DATA_BLOCK "DB LAUER"
TITLE =
VERSION : 0.0


  STRUCT
   D_0 : WORD ;
   D_1 : WORD ;
   D_2 : WORD ;
   D_3 : WORD  := W#16#A1;
   D_4 : WORD ;
   D_5 : WORD ;
   D_6 : WORD ;
   D_7 : WORD ;
   D_8 : WORD ;
   D_9 : WORD  := W#16#2006;
   D_10 : WORD  := W#16#1023;
   D_11 : WORD  := W#16#13;
   D_12 : WORD  := W#16#3439;
   D_13 : WORD  := W#16#3500;
   D_14 : WORD ;
   D_15 : WORD  := W#16#1A0;
   D_16 : WORD ;
   D_17 : WORD ;
   D_18 : WORD  := W#16#7C02;
   D_19 : WORD ;
   D_20 : WORD ;
   D_21 : WORD ;
   D_22 : WORD ;
   D_23 : WORD ;
   D_24 : WORD  := W#16#8480;
   D_25 : WORD ;
   D_26 : WORD ;
   D_27 : WORD ;
   D_28 : WORD ;
   D_29 : WORD ;
   D_30 : WORD ;
   D_31 : WORD ;
   D_32 : WORD ;
   D_33 : WORD ;
   D_34 : WORD ;
   D_35 : WORD ;
   D_36 : WORD  := W#16#F00;
   D_37 : WORD  := W#16#3001;
   D_38 : WORD ;
   D_39 : WORD ;
   D_40 : WORD ;
   D_41 : WORD ;
   D_42 : WORD ;
   D_43 : WORD ;
   D_44 : WORD ;
   D_45 : WORD ;
   D_46 : WORD ;
   D_47 : WORD ;
   D_48 : WORD ;
   D_49 : WORD ;
   D_50 : WORD ;
   D_51 : WORD ;
   D_52 : WORD ;
   D_53 : WORD ;
   D_54 : WORD ;
   D_55 : WORD ;
   D_56 : WORD ;
   D_57 : WORD ;
   D_58 : WORD ;
   D_59 : WORD ;
   D_60 : WORD ;
   D_61 : WORD ;
   D_62 : WORD ;
   D_63 : WORD ;
   D_64 : WORD ;
   D_65 : WORD ;
   D_66 : WORD ;
   D_67 : WORD ;
   D_68 : WORD ;
   D_69 : WORD ;
   D_70 : WORD ;
   D_71 : WORD ;
   D_72 : WORD ;
   D_73 : WORD ;
   D_74 : WORD ;
   D_75 : WORD ;
   D_76 : WORD ;
   D_77 : WORD  := W#16#4;
   D_78 : WORD  := W#16#2;
   D_79 : WORD  := W#16#1;
   D_80 : WORD  := W#16#1;
   D_81 : WORD  := W#16#1;
   D_82 : WORD  := W#16#1;
   D_83 : WORD  := W#16#1;
   D_84 : WORD  := W#16#2;
   D_85 : WORD  := W#16#3;
   D_86 : WORD  := W#16#2;
   D_87 : WORD  := W#16#1;
   D_88 : WORD  := W#16#1;
   D_89 : WORD  := W#16#3;
   D_90 : WORD  := W#16#4;
   D_91 : WORD  := W#16#7;
   D_92 : WORD  := W#16#9;
   D_93 : WORD  := W#16#3;
   D_94 : WORD  := W#16#3;
   D_95 : WORD  := W#16#4;
   D_96 : WORD  := W#16#1;
   D_97 : WORD  := W#16#1;
   D_98 : WORD  := W#16#1;
   D_99 : WORD  := W#16#1;
   D_100 : WORD  := W#16#1;
   D_101 : WORD  := W#16#1;
   D_102 : WORD  := W#16#1;
   D_103 : WORD ;
   D_104 : WORD ;
   D_105 : WORD ;
   D_106 : WORD ;
   D_107 : WORD ;
   D_108 : WORD ;
   D_109 : WORD ;
   D_110 : WORD  := W#16#2;
   D_111 : WORD ;
   D_112 : WORD ;
   D_113 : WORD ;
   D_114 : WORD ;
   D_115 : WORD ;
   D_116 : WORD ;
   D_117 : WORD  := W#16#7;
   D_118 : WORD  := W#16#1;
   D_119 : WORD  := W#16#1;
   D_120 : WORD  := W#16#2010;
   D_121 : WORD  := W#16#58;
   D_122 : WORD  := W#16#2010;
   D_123 : WORD  := W#16#2090;
   D_124 : WORD  := W#16#9;
   D_125 : WORD ;
   D_126 : WORD  := W#16#15;
   D_127 : WORD ;
   D_128 : WORD ;
   D_129 : WORD  := W#16#6;
   D_130 : WORD  := W#16#320;
   D_131 : WORD ;
   D_132 : WORD  := W#16#B7;
   D_133 : WORD  := W#16#1EDE;
   D_134 : WORD ;
   D_135 : WORD ;
   D_136 : WORD ;
   D_137 : WORD ;
   D_138 : WORD ;
   D_139 : WORD ;
   D_140 : WORD  := W#16#320;
   D_141 : WORD ;
   D_142 : WORD  := W#16#37;
   D_143 : WORD  := W#16#5D2;
   D_144 : WORD ;
   D_145 : WORD ;
   D_146 : WORD ;
   D_147 : WORD ;
   D_148 : WORD ;
   D_149 : WORD ;
   D_150 : WORD  := W#16#5C;
   D_151 : WORD ;
   D_152 : WORD ;
   D_153 : WORD ;
   D_154 : WORD ;
   D_155 : WORD ;
   D_156 : WORD ;
   D_157 : WORD ;
   D_158 : WORD ;
   D_159 : WORD ;
   D_160 : WORD  := W#16#320;
   D_161 : WORD ;
   D_162 : WORD  := W#16#B9;
   D_163 : WORD  := W#16#181F;
   D_164 : WORD ;
   D_165 : WORD ;
   D_166 : WORD ;
   D_167 : WORD ;
   D_168 : WORD ;
   D_169 : WORD ;
   D_170 : WORD  := W#16#320;
   D_171 : WORD ;
   D_172 : WORD  := W#16#F;
   D_173 : WORD  := W#16#14B9;
   D_174 : WORD ;
   D_175 : WORD ;
   D_176 : WORD ;
   D_177 : WORD ;
   D_178 : WORD ;
   D_179 : WORD ;
   D_180 : WORD  := W#16#320;
   D_181 : WORD ;
   D_182 : WORD ;
   D_183 : WORD  := W#16#4B0;
   D_184 : WORD  := W#16#1;
   D_185 : WORD  := W#16#1;
   D_186 : WORD ;
   D_187 : WORD ;
   D_188 : WORD ;
   D_189 : WORD ;
   D_190 : WORD ;
   D_191 : WORD ;
   D_192 : WORD ;
   D_193 : WORD ;
   D_194 : WORD ;
   D_195 : WORD ;
   D_196 : WORD ;
   D_197 : WORD ;
   D_198 : WORD ;
   D_199 : WORD ;
   D_200 : WORD ;
   D_201 : WORD ;
   D_202 : WORD ;
   D_203 : WORD ;
   D_204 : WORD ;
   D_205 : WORD ;
   D_206 : WORD ;
   D_207 : WORD ;
   D_208 : WORD ;
   D_209 : WORD ;
   D_210 : WORD ;
   D_211 : WORD ;
   D_212 : WORD ;
   D_213 : WORD ;
   D_214 : WORD ;
   D_215 : WORD ;
   D_216 : WORD ;
   D_217 : WORD ;
   D_218 : WORD ;
   D_219 : WORD ;
   D_220 : WORD ;
   D_221 : WORD ;
   D_222 : WORD ;
   D_223 : WORD ;
   D_224 : WORD ;
   D_225 : WORD ;
   D_226 : WORD ;
   D_227 : WORD ;
   D_228 : WORD ;
   D_229 : WORD ;
   D_230 : WORD ;
   D_231 : WORD ;
   D_232 : WORD ;
   D_233 : WORD ;
   D_234 : WORD ;
   D_235 : WORD ;
   D_236 : WORD ;
   D_237 : WORD ;
   D_238 : WORD ;
   D_239 : WORD ;
   D_240 : WORD ;
   D_241 : WORD ;
   D_242 : WORD ;
   D_243 : WORD ;
   D_244 : WORD ;
   D_245 : WORD ;
   D_246 : WORD ;
   D_247 : WORD ;
   D_248 : WORD ;
   D_249 : WORD ;
   D_250 : WORD ;
   D_251 : WORD ;
   D_252 : WORD  := W#16#58;
   D_253 : WORD  := W#16#9;
   D_254 : WORD ;
   D_255 : WORD  := W#16#12;
  END_STRUCT ;
BEGIN
   D_0 := W#16#4B;
   D_1 := W#16#0;
   D_2 := W#16#0;
   D_3 := W#16#0;
   D_4 := W#16#0;
   D_5 := W#16#0;
   D_6 := W#16#0;
   D_7 := W#16#0;
   D_8 := W#16#0;
   D_9 := W#16#2010;
   D_10 := W#16#527;
   D_11 := W#16#619;
   D_12 := W#16#306;
   D_13 := W#16#3F00;
   D_14 := W#16#0;
   D_15 := W#16#1A0;
   D_16 := W#16#0;
   D_17 := W#16#0;
   D_18 := W#16#7C02;
   D_19 := W#16#0;
   D_20 := W#16#0;
   D_21 := W#16#0;
   D_22 := W#16#0;
   D_23 := W#16#0;
   D_24 := W#16#8480;
   D_25 := W#16#0;
   D_26 := W#16#0;
   D_27 := W#16#0;
   D_28 := W#16#0;
   D_29 := W#16#0;
   D_30 := W#16#0;
   D_31 := W#16#0;
   D_32 := W#16#0;
   D_33 := W#16#0;
   D_34 := W#16#0;
   D_35 := W#16#0;
   D_36 := W#16#F00;
   D_37 := W#16#3001;
   D_38 := W#16#0;
   D_39 := W#16#0;
   D_40 := W#16#0;
   D_41 := W#16#0;
   D_42 := W#16#0;
   D_43 := W#16#0;
   D_44 := W#16#0;
   D_45 := W#16#0;
   D_46 := W#16#0;
   D_47 := W#16#0;
   D_48 := W#16#0;
   D_49 := W#16#0;
   D_50 := W#16#0;
   D_51 := W#16#0;
   D_52 := W#16#0;
   D_53 := W#16#0;
   D_54 := W#16#0;
   D_55 := W#16#0;
   D_56 := W#16#0;
   D_57 := W#16#0;
   D_58 := W#16#0;
   D_59 := W#16#0;
   D_60 := W#16#0;
   D_61 := W#16#0;
   D_62 := W#16#0;
   D_63 := W#16#0;
   D_64 := W#16#0;
   D_65 := W#16#0;
   D_66 := W#16#0;
   D_67 := W#16#0;
   D_68 := W#16#0;
   D_69 := W#16#0;
   D_70 := W#16#0;
   D_71 := W#16#0;
   D_72 := W#16#0;
   D_73 := W#16#0;
   D_74 := W#16#0;
   D_75 := W#16#0;
   D_76 := W#16#0;
   D_77 := W#16#4;
   D_78 := W#16#2;
   D_79 := W#16#4;
   D_80 := W#16#1;
   D_81 := W#16#1;
   D_82 := W#16#1;
   D_83 := W#16#1;
   D_84 := W#16#A;
   D_85 := W#16#4;
   D_86 := W#16#9;
   D_87 := W#16#1;
   D_88 := W#16#1;
   D_89 := W#16#1;
   D_90 := W#16#4;
   D_91 := W#16#7;
   D_92 := W#16#9;
   D_93 := W#16#4;
   D_94 := W#16#2;
   D_95 := W#16#1;
   D_96 := W#16#0;
   D_97 := W#16#0;
   D_98 := W#16#0;
   D_99 := W#16#0;
   D_100 := W#16#0;
   D_101 := W#16#1;
   D_102 := W#16#0;
   D_103 := W#16#0;
   D_104 := W#16#0;
   D_105 := W#16#0;
   D_106 := W#16#0;
   D_107 := W#16#0;
   D_108 := W#16#0;
   D_109 := W#16#0;
   D_110 := W#16#2;
   D_111 := W#16#0;
   D_112 := W#16#0;
   D_113 := W#16#0;
   D_114 := W#16#C;
   D_115 := W#16#C;
   D_116 := W#16#1;
   D_117 := W#16#7;
   D_118 := W#16#0;
   D_119 := W#16#1;
   D_120 := W#16#2010;
   D_121 := W#16#96;
   D_122 := W#16#2010;
   D_123 := W#16#2090;
   D_124 := W#16#C;
   D_125 := W#16#0;
   D_126 := W#16#15;
   D_127 := W#16#0;
   D_128 := W#16#0;
   D_129 := W#16#6;
   D_130 := W#16#320;
   D_131 := W#16#0;
   D_132 := W#16#2A9;
   D_133 := W#16#238;
   D_134 := W#16#0;
   D_135 := W#16#0;
   D_136 := W#16#0;
   D_137 := W#16#0;
   D_138 := W#16#0;
   D_139 := W#16#0;
   D_140 := W#16#320;
   D_141 := W#16#0;
   D_142 := W#16#98;
   D_143 := W#16#1262;
   D_144 := W#16#0;
   D_145 := W#16#0;
   D_146 := W#16#0;
   D_147 := W#16#0;
   D_148 := W#16#0;
   D_149 := W#16#0;
   D_150 := W#16#67;
   D_151 := W#16#0;
   D_152 := W#16#0;
   D_153 := W#16#0;
   D_154 := W#16#0;
   D_155 := W#16#0;
   D_156 := W#16#0;
   D_157 := W#16#0;
   D_158 := W#16#0;
   D_159 := W#16#0;
   D_160 := W#16#320;
   D_161 := W#16#0;
   D_162 := W#16#2C1;
   D_163 := W#16#FD0;
   D_164 := W#16#0;
   D_165 := W#16#0;
   D_166 := W#16#0;
   D_167 := W#16#0;
   D_168 := W#16#0;
   D_169 := W#16#0;
   D_170 := W#16#320;
   D_171 := W#16#0;
   D_172 := W#16#0;
   D_173 := W#16#0;
   D_174 := W#16#1;
   D_175 := W#16#1;
   D_176 := W#16#0;
   D_177 := W#16#0;
   D_178 := W#16#0;
   D_179 := W#16#0;
   D_180 := W#16#320;
   D_181 := W#16#0;
   D_182 := W#16#0;
   D_183 := W#16#7B0;
   D_184 := W#16#1;
   D_185 := W#16#1;
   D_186 := W#16#0;
   D_187 := W#16#0;
   D_188 := W#16#0;
   D_189 := W#16#0;
   D_190 := W#16#0;
   D_191 := W#16#0;
   D_192 := W#16#0;
   D_193 := W#16#0;
   D_194 := W#16#0;
   D_195 := W#16#0;
   D_196 := W#16#0;
   D_197 := W#16#0;
   D_198 := W#16#0;
   D_199 := W#16#0;
   D_200 := W#16#0;
   D_201 := W#16#0;
   D_202 := W#16#0;
   D_203 := W#16#0;
   D_204 := W#16#0;
   D_205 := W#16#0;
   D_206 := W#16#0;
   D_207 := W#16#0;
   D_208 := W#16#0;
   D_209 := W#16#0;
   D_210 := W#16#0;
   D_211 := W#16#0;
   D_212 := W#16#0;
   D_213 := W#16#0;
   D_214 := W#16#0;
   D_215 := W#16#0;
   D_216 := W#16#0;
   D_217 := W#16#0;
   D_218 := W#16#0;
   D_219 := W#16#0;
   D_220 := W#16#0;
   D_221 := W#16#0;
   D_222 := W#16#0;
   D_223 := W#16#0;
   D_224 := W#16#0;
   D_225 := W#16#0;
   D_226 := W#16#0;
   D_227 := W#16#0;
   D_228 := W#16#0;
   D_229 := W#16#0;
   D_230 := W#16#0;
   D_231 := W#16#0;
   D_232 := W#16#0;
   D_233 := W#16#0;
   D_234 := W#16#0;
   D_235 := W#16#0;
   D_236 := W#16#0;
   D_237 := W#16#0;
   D_238 := W#16#0;
   D_239 := W#16#0;
   D_240 := W#16#0;
   D_241 := W#16#0;
   D_242 := W#16#0;
   D_243 := W#16#0;
   D_244 := W#16#0;
   D_245 := W#16#0;
   D_246 := W#16#0;
   D_247 := W#16#0;
   D_248 := W#16#0;
   D_249 := W#16#0;
   D_250 := W#16#0;
   D_251 := W#16#0;
   D_252 := W#16#C;
   D_253 := W#16#12;
   D_254 := W#16#0;
   D_255 := W#16#12;
END_DATA_BLOCK
